(* CODESYS project visu_iol_o5d150_v1.export

Project tree, tasks and I/O mapping:
  visualisation Visu_IOL_O5D150
*)

// /Visu_IOL_O5D150
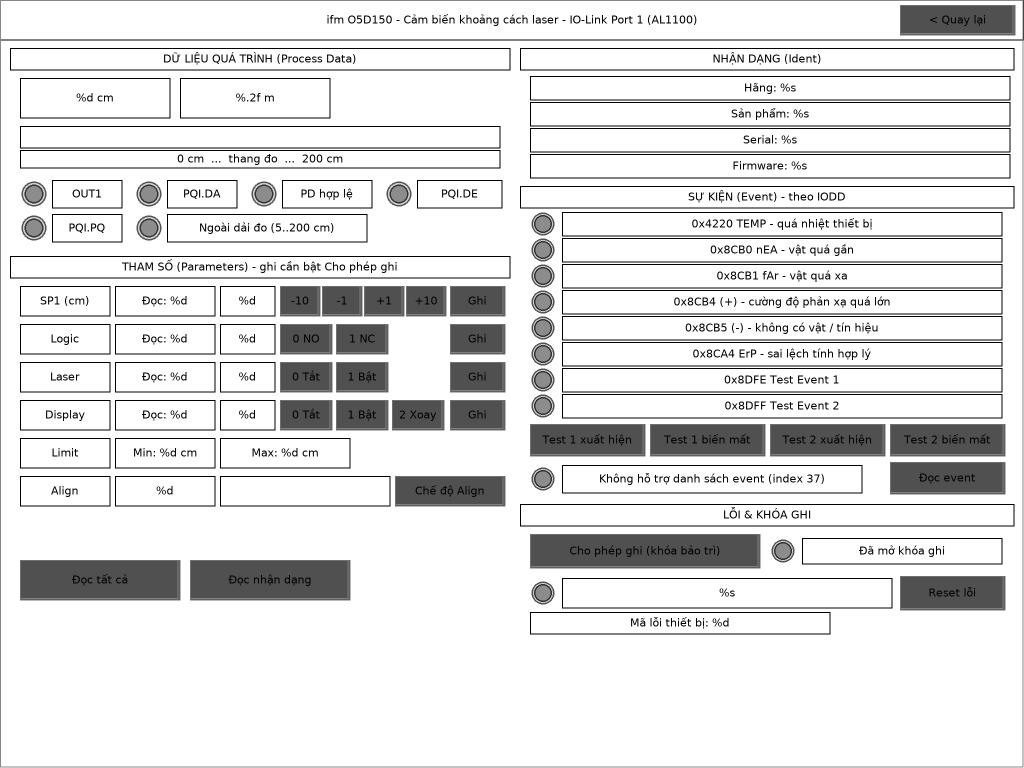
VISUALIZATION Visu_IOL_O5D150  // 1024x768
    Rectangle (0,0 1024x40), "ifm O5D150 - Cảm biến khoảng cách laser - IO-Link Port 1 (AL1100)"
    Button (900,5 115x30), "< Quay lại"
        OnMouseClick:  Assign=Visu_Main, Type=Assignment
    Rectangle (10,48 500x22), "DỮ LIỆU QUÁ TRÌNH (Process Data)"
    Rectangle (20,78 150x40), "%d cm", text variable: GVL_HMI_IOL.stO5D150.uiDistance_cm
    Rectangle (180,78 150x40), "%.2f m", text variable: GVL_HMI_IOL.stO5D150.rDistance_m
    Rectangle (20,126 480x22)
    Rectangle (20,126 480x22)
        p874137650: -(480 - MIN(480, UINT_TO_INT(GVL_HMI_IOL.stO5D150.uiDistance_cm) * 480 / 200))
    Rectangle (20,150 480x18), "0 cm ... thang đo ... 200 cm"
    Lamp1 (20,180 28x28), variable: GVL_HMI_IOL.stO5D150.xOut1, style: Lamp-Lamp1-Gray
    Rectangle (52,180 70x28), "OUT1"
    Lamp1 (135,180 28x28), variable: GVL_HMI_IOL.stO5D150.xDA, style: Lamp-Lamp1-Gray
    Rectangle (167,180 70x28), "PQI.DA"
    Lamp1 (250,180 28x28), variable: GVL_HMI_IOL.stO5D150.xPdValid, style: Lamp-Lamp1-Gray
    Rectangle (282,180 90x28), "PD hợp lệ"
    Lamp1 (385,180 28x28), variable: GVL_HMI_IOL.stO5D150.xDE, style: Lamp-Lamp1-Gray
    Rectangle (417,180 85x28), "PQI.DE"
    Lamp1 (20,214 28x28), variable: GVL_HMI_IOL.stO5D150.xPQ, style: Lamp-Lamp1-Gray
    Rectangle (52,214 70x28), "PQI.PQ"
    Lamp1 (135,214 28x28), variable: GVL_HMI_IOL.stO5D150.xOutOfRange, style: Lamp-Lamp1-Gray
    Rectangle (167,214 200x28), "Ngoài dải đo (5..200 cm)"
    Rectangle (10,256 500x22), "THAM SỐ (Parameters) - ghi cần bật Cho phép ghi"
    Rectangle (20,286 90x30), "SP1 (cm)"
    Rectangle (115,286 100x30), "Đọc: %d", text variable: GVL_HMI_IOL.stO5D150.uiSP1
    Rectangle (220,286 55x30), "%d", text variable: GVL_HMI_IOL.stO5D150.uiSetSP1
    Button (280,286 40x30), "-10", input disabled if: NOT GVL_HMI_IOL.xMaintEnable
        OnMouseClick: execute { GVL_HMI_IOL.stO5D150.uiSetSP1 := DINT_TO_UINT(LIMIT(5, UINT_TO_DINT(GVL_HMI_IOL.stO5D150.uiSetSP1) + (-10), 200)); }
    Button (322,286 40x30), "-1", input disabled if: NOT GVL_HMI_IOL.xMaintEnable
        OnMouseClick: execute { GVL_HMI_IOL.stO5D150.uiSetSP1 := DINT_TO_UINT(LIMIT(5, UINT_TO_DINT(GVL_HMI_IOL.stO5D150.uiSetSP1) + (-1), 200)); }
    Button (364,286 40x30), "+1", input disabled if: NOT GVL_HMI_IOL.xMaintEnable
        OnMouseClick: execute { GVL_HMI_IOL.stO5D150.uiSetSP1 := DINT_TO_UINT(LIMIT(5, UINT_TO_DINT(GVL_HMI_IOL.stO5D150.uiSetSP1) + (1), 200)); }
    Button (406,286 40x30), "+10", input disabled if: NOT GVL_HMI_IOL.xMaintEnable
        OnMouseClick: execute { GVL_HMI_IOL.stO5D150.uiSetSP1 := DINT_TO_UINT(LIMIT(5, UINT_TO_DINT(GVL_HMI_IOL.stO5D150.uiSetSP1) + (10), 200)); }
    Button (450,286 55x30), "Ghi", input disabled if: NOT GVL_HMI_IOL.xMaintEnable
        OnMouseClick: execute { GVL_HMI_IOL.stO5D150.xCmdWriteSP1 := TRUE; }
    Rectangle (20,324 90x30), "Logic"
    Rectangle (115,324 100x30), "Đọc: %d", text variable: GVL_HMI_IOL.stO5D150.usiLogic
    Rectangle (220,324 55x30), "%d", text variable: GVL_HMI_IOL.stO5D150.usiSetLogic
    Button (280,324 52x30), "0 NO", input disabled if: NOT GVL_HMI_IOL.xMaintEnable
        OnMouseClick: execute { GVL_HMI_IOL.stO5D150.usiSetLogic := 0; }
    Button (336,324 52x30), "1 NC", input disabled if: NOT GVL_HMI_IOL.xMaintEnable
        OnMouseClick: execute { GVL_HMI_IOL.stO5D150.usiSetLogic := 1; }
    Button (450,324 55x30), "Ghi", input disabled if: NOT GVL_HMI_IOL.xMaintEnable
        OnMouseClick: execute { GVL_HMI_IOL.stO5D150.xCmdWriteLogic := TRUE; }
    Rectangle (20,362 90x30), "Laser"
    Rectangle (115,362 100x30), "Đọc: %d", text variable: GVL_HMI_IOL.stO5D150.usiLaser
    Rectangle (220,362 55x30), "%d", text variable: GVL_HMI_IOL.stO5D150.usiSetLaser
    Button (280,362 52x30), "0 Tắt", input disabled if: NOT GVL_HMI_IOL.xMaintEnable
        OnMouseClick: execute { GVL_HMI_IOL.stO5D150.usiSetLaser := 0; }
    Button (336,362 52x30), "1 Bật", input disabled if: NOT GVL_HMI_IOL.xMaintEnable
        OnMouseClick: execute { GVL_HMI_IOL.stO5D150.usiSetLaser := 1; }
    Button (450,362 55x30), "Ghi", input disabled if: NOT GVL_HMI_IOL.xMaintEnable
        OnMouseClick: execute { GVL_HMI_IOL.stO5D150.xCmdWriteLaser := TRUE; }
    Rectangle (20,400 90x30), "Display"
    Rectangle (115,400 100x30), "Đọc: %d", text variable: GVL_HMI_IOL.stO5D150.usiDisplay
    Rectangle (220,400 55x30), "%d", text variable: GVL_HMI_IOL.stO5D150.usiSetDisplay
    Button (280,400 52x30), "0 Tắt", input disabled if: NOT GVL_HMI_IOL.xMaintEnable
        OnMouseClick: execute { GVL_HMI_IOL.stO5D150.usiSetDisplay := 0; }
    Button (336,400 52x30), "1 Bật", input disabled if: NOT GVL_HMI_IOL.xMaintEnable
        OnMouseClick: execute { GVL_HMI_IOL.stO5D150.usiSetDisplay := 1; }
    Button (392,400 52x30), "2 Xoay", input disabled if: NOT GVL_HMI_IOL.xMaintEnable
        OnMouseClick: execute { GVL_HMI_IOL.stO5D150.usiSetDisplay := 2; }
    Button (450,400 55x30), "Ghi", input disabled if: NOT GVL_HMI_IOL.xMaintEnable
        OnMouseClick: execute { GVL_HMI_IOL.stO5D150.xCmdWriteDisplay := TRUE; }
    Rectangle (20,438 90x30), "Limit"
    Rectangle (115,438 100x30), "Min: %d cm", text variable: GVL_HMI_IOL.stO5D150.uiLimitMin_cm
    Rectangle (220,438 130x30), "Max: %d cm", text variable: GVL_HMI_IOL.stO5D150.uiLimitMax_cm
    Rectangle (20,476 90x30), "Align"
    Rectangle (115,476 100x30), "%d", text variable: GVL_HMI_IOL.stO5D150.usiAlign
    Rectangle (220,476 170x30)
    Rectangle (220,476 170x30)
        p874137650: -(170 - MIN(170, USINT_TO_INT(GVL_HMI_IOL.stO5D150.usiAlign) * 170 / 100))
    Button (395,476 110x30), "Chế độ Align"
        OnMouseClick: execute { GVL_HMI_IOL.stO5D150.xAlignMode := NOT GVL_HMI_IOL.stO5D150.xAlignMode; }
    Button (20,560 160x40), "Đọc tất cả"
        OnMouseClick: execute { GVL_HMI_IOL.stO5D150.xCmdReadAll := TRUE; }
    Button (190,560 160x40), "Đọc nhận dạng"
        OnMouseClick: execute { GVL_HMI_IOL.stO5D150.xCmdReadIdent := TRUE; }
    Rectangle (520,48 494x22), "NHẬN DẠNG (Ident)"
    Rectangle (530,76 480x24), "Hãng: %s", text variable: GVL_HMI_IOL.stO5D150.sVendor
    Rectangle (530,102 480x24), "Sản phẩm: %s", text variable: GVL_HMI_IOL.stO5D150.sProduct
    Rectangle (530,128 480x24), "Serial: %s", text variable: GVL_HMI_IOL.stO5D150.sSerial
    Rectangle (530,154 480x24), "Firmware: %s", text variable: GVL_HMI_IOL.stO5D150.sFwRev
    Rectangle (520,186 494x22), "SỰ KIỆN (Event) - theo IODD"
    Lamp1 (530,211 26x26), variable: GVL_HMI_IOL.stO5D150.axEvtActive[0], style: Lamp-Lamp1-Gray
    Rectangle (562,212 440x24), "0x4220 TEMP - quá nhiệt thiết bị"
    Lamp1 (530,237 26x26), variable: GVL_HMI_IOL.stO5D150.axEvtActive[1], style: Lamp-Lamp1-Gray
    Rectangle (562,238 440x24), "0x8CB0 nEA - vật quá gần"
    Lamp1 (530,263 26x26), variable: GVL_HMI_IOL.stO5D150.axEvtActive[2], style: Lamp-Lamp1-Gray
    Rectangle (562,264 440x24), "0x8CB1 fAr - vật quá xa"
    Lamp1 (530,289 26x26), variable: GVL_HMI_IOL.stO5D150.axEvtActive[3], style: Lamp-Lamp1-Gray
    Rectangle (562,290 440x24), "0x8CB4 (+) - cường độ phản xạ quá lớn"
    Lamp1 (530,315 26x26), variable: GVL_HMI_IOL.stO5D150.axEvtActive[4], style: Lamp-Lamp1-Gray
    Rectangle (562,316 440x24), "0x8CB5 (-) - không có vật / tín hiệu"
    Lamp1 (530,341 26x26), variable: GVL_HMI_IOL.stO5D150.axEvtActive[5], style: Lamp-Lamp1-Gray
    Rectangle (562,342 440x24), "0x8CA4 ErP - sai lệch tính hợp lý"
    Lamp1 (530,367 26x26), variable: GVL_HMI_IOL.stO5D150.axEvtActive[6], style: Lamp-Lamp1-Gray
    Rectangle (562,368 440x24), "0x8DFE Test Event 1"
    Lamp1 (530,393 26x26), variable: GVL_HMI_IOL.stO5D150.axEvtActive[7], style: Lamp-Lamp1-Gray
    Rectangle (562,394 440x24), "0x8DFF Test Event 2"
    Button (530,424 115x32), "Test 1 xuất hiện", input disabled if: NOT GVL_HMI_IOL.xMaintEnable
        OnMouseClick: execute { GVL_HMI_IOL.stO5D150.xCmdTestEvt1On := TRUE; }
    Button (650,424 115x32), "Test 1 biến mất", input disabled if: NOT GVL_HMI_IOL.xMaintEnable
        OnMouseClick: execute { GVL_HMI_IOL.stO5D150.xCmdTestEvt1Off := TRUE; }
    Button (770,424 115x32), "Test 2 xuất hiện", input disabled if: NOT GVL_HMI_IOL.xMaintEnable
        OnMouseClick: execute { GVL_HMI_IOL.stO5D150.xCmdTestEvt2On := TRUE; }
    Button (890,424 115x32), "Test 2 biến mất", input disabled if: NOT GVL_HMI_IOL.xMaintEnable
        OnMouseClick: execute { GVL_HMI_IOL.stO5D150.xCmdTestEvt2Off := TRUE; }
    Lamp1 (530,466 26x26), variable: GVL_HMI_IOL.stO5D150.xEvtListNotSupported, style: Lamp-Lamp1-Gray
    Rectangle (562,465 300x28), "Không hỗ trợ danh sách event (index 37)"
    Button (890,462 115x32), "Đọc event"
        OnMouseClick: execute { GVL_HMI_IOL.stO5D150.xCmdReadEvents := TRUE; }
    Rectangle (520,504 494x22), "LỖI & KHÓA GHI"
    Button (530,534 230x34), "Cho phép ghi (khóa bảo trì)"
        OnMouseClick: execute { GVL_HMI_IOL.xMaintEnable := NOT GVL_HMI_IOL.xMaintEnable; }
    Lamp1 (770,538 26x26), variable: GVL_HMI_IOL.xMaintEnable, style: Lamp-Lamp1-Gray
    Rectangle (802,538 200x26), "Đã mở khóa ghi"
    Lamp1 (530,580 26x26), variable: GVL_HMI_IOL.stO5D150.xError, style: Lamp-Lamp1-Gray
    Rectangle (562,578 330x30), "%s", text variable: GVL_HMI_IOL.stO5D150.wsErrText
    Button (900,576 105x34), "Reset lỗi"
        OnMouseClick: execute { GVL_HMI_IOL.stO5D150.xCmdResetErr := TRUE; }
    Rectangle (530,612 300x22), "Mã lỗi thiết bị: %d", text variable: GVL_HMI_IOL.stO5D150.uiDevErr
END_VISUALIZATION
